TYPE U_MOVER_SELECTOR_STATE :
UNION
  stState             : ST_MOVER_SELECTOR_STATE;

  byState   AT %I*    : ARRAY[1..SIZEOF(ST_MOVER_SELECTOR_STATE)] OF BYTE;
END_UNION
END_TYPE

(* stored: Version 1.1.0.1
   DUT U_MOVER_SELECTOR_STATE: Id {5ebf3bd4-1a93-4353-b1e5-ab3be2d85495} *)
